(* PLC project marcha_paro, UCuenca DEET Tablero DEET 1 *)
(* stored: creationDateTime 2026-10-19T12:00:00, modificationDateTime 2026-10-19T12:00:00 *)

(* Marcha/paro con enclavamiento: I16 arranca D18, I18 lo para. *)
PROGRAM marcha_paro
  VAR
    MARCHA AT %IX102.0 : BOOL;  (* Pulsador I16 del Controllino *)
    PARO AT %IX102.2 : BOOL;  (* Pulsador I18 del Controllino *)
    MOTOR AT %QX102.2 : BOOL;  (* Salida D18 del Controllino *)
  END_VAR

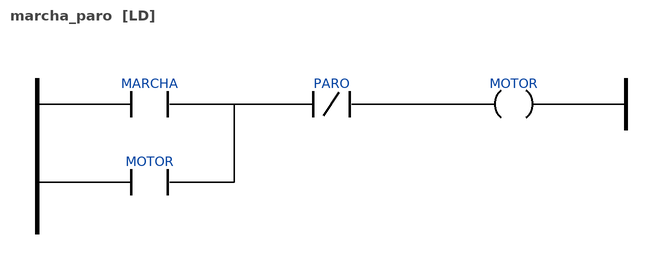
(* LD diagram, written out as Structured Text *)
MOTOR := (MARCHA OR MOTOR) AND NOT PARO;
END_PROGRAM

CONFIGURATION Config0
  RESOURCE Res0 ON PLC
    TASK task0(INTERVAL := T#20ms, PRIORITY := 0);
    PROGRAM instance0 WITH task0 : marcha_paro;
  END_RESOURCE
END_CONFIGURATION
